(* IEC 61131-3 sources: Masterarbeit/sigmatek/lasalclass2/PW022_virtualization/Network, 1 file *)

(* ---- ConfigObjects.st ---- *)
FUNCTION GLOBAL TAB TASK_CONF
_K_TASK, _K_REAL,
_K_END_VAR,

_K_TASK, _K_CYCLIC,
_K_END_VAR,

_K_TASK, _K_BACKGROUND,
_K_END_VAR,

_K_END_CONF
END_FUNCTION

FUNCTION GLOBAL TAB IPR_CONF
_K_IPR
	0$UINT,
_K_END_VAR,
_K_END_CONF
END_FUNCTION

FUNCTION GLOBAL TAB CONFIG_TABLES
00063$UINT,
0$UINT, 1, 14, "_BUSINTERFACESDIASDRIVEMNG",
0$UINT, 0, 4, "_CAN",
0$UINT, 1, 10, "_CANLIB",
0$UINT, 1, 72, "_DRIVEAXIS",
0$UINT, 1, 81, "_DRIVEAXISBASE",
0$UINT, 1, 22, "_DRIVEAXISSET",
0$UINT, 1, 82, "_DRIVEMNG_DC062",
0$UINT, 1, 61, "_DRIVEMNGBASE",
0$UINT, 1, 20, "_FILESYS",
0$UINT, 0, 5, "_LINKER",
0$UINT, 1, 3, "_LOADSIMULATOR",
0$UINT, 1, 1, "_MULTITASK",
0$UINT, 0, 5, "_OSKERNEL",
0$UINT, 1, 34, "_SERLIB",
0$UINT, 0, 0, "_STDLIB",
0$UINT, 1, 1, "_TASKOBJECTCONTROL",
0$UINT, 1, 69, "_VARANDRIVEBASE",
0$UINT, 1, 38, "AO081",
0$UINT, 1, 21, "ASCII_BIN",
0$UINT, 2, 1, "BUSINTERFACESDIASINTERNAL",
0$UINT, 1, 75, "BUSINTERFACEVARAN",
0$UINT, 1, 2, "CP841_IOS",
0$UINT, 0, 4, "CRITICALSECTION",
0$UINT, 2, 33, "DIASMASTER",
0$UINT, 1, 83, "DIASMASTERC",
0$UINT, 2, 25, "DIASMASTERMAIN",
0$UINT, 1, 0, "DIASMASTERPOSTSCAN",
0$UINT, 1, 13, "DM081",
0$UINT, 1, 11, "EEPROM",
0$UINT, 1, 21, "HUB_BASE",
0$UINT, 2, 11, "HUB_BASE_ROOT",
0$UINT, 2, 36, "HWBASE",
0$UINT, 2, 56, "HWBASECDIAS",
0$UINT, 1, 0, "HWCLOGGING",
0$UINT, 5, 21, "HWCONTROL",
0$UINT, 1, 10, "HWCONTROLBASE",
0$UINT, 1, 0, "HWRTPOSTSCAN",
0$UINT, 1, 6, "I2CCDIAS",
0$UINT, 1, 22, "MERKEREX",
0$UINT, 1, 5, "PW022",
0$UINT, 1, 17, "RAMEX",
0$UINT, 1, 9, "RAMFILE",
0$UINT, 3, 19, "SAFETYCDIAS_BASE",
0$UINT, 2, 26, "SAFETYMANAGER",
0$UINT, 1, 4, "SAFETYUDP",
0$UINT, 1, 60, "SDIASBASE",
0$UINT, 1, 10, "SDIASHUBBASE",
0$UINT, 1, 97, "SDIASMANAGER",
0$UINT, 2, 6, "SDIASPLC",
0$UINT, 0, 41, "SIGCLIB",
0$UINT, 0, 0, "STEUERUNG",
0$UINT, 1, 11, "STRING",
0$UINT, 1, 85, "STRINGINTERNAL",
0$UINT, 1, 21, "SYNCCALL",
0$UINT, 2, 20, "VARAN_BASE",
0$UINT, 3, 7, "VARANMANAGER",
0$UINT, 2, 7, "VARANMANAGER_1",
0$UINT, 2, 9, "VARANMANAGER_2",
0$UINT, 1, 26, "VARANMANAGER_BASE",
0$UINT, 1, 101, "VI021",
0$UINT, 1, 3, "VIRTUALBASEINIT",
0$UINT, 2, 11, "WATCHDOGDIAS",
0$UINT, 1, 1, "XXXBASE_IOS",
ONE_CFG$UINT, 0, 0, "ONE_HW_Network",
TASK_CFG$UINT, 0, 0, "TASK_CONF",
IPR_CFG$UINT, 0, 0, "IPR_CONF",
PRJ_CFG$UINT, 0, 0, "PW022_virtualization",
END_FUNCTION

#ifdef __LSLLDR_IOELEMENTS__
FUNCTION GLOBAL TAB _IO_ELEMENTS_TAB
0001$UINT, 0001$UINT,
"**IOCONN_EMPTY**", "PW022_1_Copy.PeriodeDuration_Ch1",
0012$UINT,
"**IOCONN_EMPTY**", "Steuerung1.cPeriodeDuration_ch3",
"**IOCONN_EMPTY**", "Steuerung1.cPeriodeDuration_ch1",
"**IOCONN_EMPTY**", "Steuerung1.cPWMOnTime_ch1",
"**IOCONN_EMPTY**", "Steuerung1.cPeriodeDuration_ch2",
"**IOCONN_EMPTY**", "Steuerung1.cPWMOnTime_ch2",
"**IOCONN_EMPTY**", "Steuerung1.cPWMOnTime_ch3",
"**IOCONN_EMPTY**", "Steuerung1.cPeriodeDuration_ch4",
"**IOCONN_EMPTY**", "Steuerung1.cPWMOnTime_ch4",
"**IOCONN_EMPTY**", "Steuerung1.cPeriodeDuration_ch5",
"**IOCONN_EMPTY**", "Steuerung1.cPWMOnTime_ch5",
"**IOCONN_EMPTY**", "Steuerung1.cPeriodeDuration_ch6",
"**IOCONN_EMPTY**", "Steuerung1.cPWMOnTime_ch6",
END_FUNCTION
#endif //__LSLLDR_IOELEMENTS__

FUNCTION GLOBAL TAB CH_REDIRECT_EMB_TAB
0000$UINT,
00015$UINT,
"_BUSINTERFACESDIASDRIVEMNG;SERIALNO", "\SERIALNOSTR.DATA",
"_DRIVEMNG_DC062;FWDATETR", "\FWDATESTRING.DATA",
"_DRIVEMNG_DC062;FWDATE", "\FWDATESTRING.DATA",
"_DRIVEMNG_DC062;FWNUMSTR", "\FWNUMSTRING.DATA",
"_DRIVEMNG_DC062;FWVERSION", "\FWNUMSTRING.DATA",
"_VARANDRIVEBASE;SERIALNO", "\SERIALNOSTR.DATA",
"AO081;SERIALNO", "\SERIALNOSTR.DATA",
"BUSINTERFACEVARAN;SERIALNO", "\SERIALNOSTR.DATA",
"DM081;SERIALNO", "\SERIALNOSTR.DATA",
"HWBASECDIAS;SERIALNO", "\SERIALNOSTR.DATA",
"PW022;SERIALNO", "\SERIALNOSTR.DATA",
"SAFETYCDIAS_BASE;SERIALNO", "\SERIALNOSTR.DATA",
"SDIASBASE;SERIALNO", "\SERIALNOSTR.DATA",
"VARAN_BASE;SERIALNO", "\SERIALNOSTR.DATA",
"VI021;SERIALNO", "\SERIALNOSTR.DATA",
END_FUNCTION
